(* IEC 61131-3 sources: plc-st-coding-agent/progress/evidence/f14_p1_20261111b/jobs/custom_minimax-m27, 44 files *)

(* ---- public-hard-01.candidate_01.st ---- *)
(* Material Proportioning Process Control *)
(* PLC Program in Structured Text (ST) *)

TYPE ProcessState :
    (
        IDLE        := 0,
        FILL_A      := 1,
        FILL_B      := 2,
        FILL_C      := 3,
        MIXING      := 4,
        DISCHARGE   := 5
    );
END_TYPE

VAR
    (* Internal state variables *)
    autoState         : ProcessState := IDLE;
    prevAutoStart     : BOOL := FALSE;
    prevValveAStart   : BOOL := FALSE;
    prevValveBStart   : BOOL := FALSE;
    prevValveCStart   : BOOL := FALSE;
    prevValveDStart   : BOOL := FALSE;
    prevMixMotorStart : BOOL := FALSE;
END_VAR

(* Emergency Stop - Highest Priority *)
IF NOT estop THEN
    valveARun    := FALSE;
    valveBRun    := FALSE;
    valveCRun    := FALSE;
    valveDRun    := FALSE;
    mixMotorRun  := FALSE;
    autoState    := IDLE;
    RETURN;
END_IF

(* Rising edge detection for buttons *)
IF autoStart AND NOT prevAutoStart THEN
    (* Rising edge detected for autoStart *)
END_IF

IF valveAStart AND NOT prevValveAStart THEN
    valveARun := NOT valveARun;
END_IF;

IF valveBStart AND NOT prevValveBStart THEN
    valveBRun := NOT valveBRun;
END_IF;

IF valveCStart AND NOT prevValveCStart THEN
    valveCRun := NOT valveCRun;
END_IF;

IF valveDStart AND NOT prevValveDStart THEN
    valveDRun := NOT valveDRun;
END_IF;

IF mixMotorStart AND NOT prevMixMotorStart THEN
    mixMotorRun := NOT mixMotorRun;
END_IF;

(* Update previous button states *)
prevAutoStart     := autoStart;
prevValveAStart   := valveAStart;
prevValveBStart   := valveBStart;
prevValveCStart   := valveCStart;
prevValveDStart   := valveDStart;
prevMixMotorStart := mixMotorStart;

(* Mode Selection *)
IF opeMode THEN
    (* ========== AUTOMATIC MODE ========== *)

    (* Initialize outputs to FALSE *)
    valveARun   := FALSE;
    valveBRun   := FALSE;
    valveCRun   := FALSE;
    valveDRun   := FALSE;
    mixMotorRun := FALSE;

    (* Start automatic process on rising edge of autoStart *)
    IF autoStart AND NOT prevAutoStart THEN
        IF autoState = IDLE THEN
            autoState := FILL_A;
            valveARun := TRUE;
        END_IF
    END_IF

    (* State Machine - Sequential Control *)
    IF autoState = FILL_A THEN
        valveARun := TRUE;
        (* When level reaches 50cm, close valve A and open valve B *)
        IF levelSensor >= 50 THEN
            autoState  := FILL_B;
            valveARun  := FALSE;
            valveBRun  := TRUE;
        END_IF

    ELSIF autoState = FILL_B THEN
        valveBRun := TRUE;
        (* When level reaches 80cm, close valve B *)
        IF levelSensor >= 80 THEN
            valveBRun := FALSE;

            (* Check processMode for next step *)
            IF NOT processMode THEN
                (* processMode=false: Direct to mixing *)
                autoState  := MIXING;
                mixMotorRun := TRUE;
            ELSE
                (* processMode=true: Fill material C first *)
                autoState := FILL_C;
            END_IF
        END_IF

    ELSIF autoState = FILL_C THEN
        valveCRun := TRUE;
        (* When level reaches 100cm, close valve C and start mixing *)
        IF levelSensor >= 100 THEN
            autoState  := MIXING;
            valveCRun  := FALSE;
            mixMotorRun := TRUE;
        END_IF

    ELSIF autoState = MIXING THEN
        mixMotorRun := TRUE;
        (* When mixing complete signal received, stop motor *)
        IF mixMotorComplete THEN
            autoState  := DISCHARGE;
            mixMotorRun := FALSE;
        END_IF

    ELSIF autoState = DISCHARGE THEN
        valveDRun := TRUE;
        (* After discharge, return to idle - process complete *)
        autoState := IDLE;

    END_IF

ELSE
    (* ========== MANUAL MODE ========== *)
    (* In manual mode, automatic state machine is reset *)
    autoState := IDLE;

END_IF

(* ---- public-medium-05.candidate_01.st ---- *)
// Automated Production Line Control - ST Implementation

// Define the states for automatic mode
TYPE ProductionState :
(
    WAIT_A           := 0,  // Waiting for product at Workstation A
    WAIT_A_PRESSED   := 1,  // Product at A, waiting for ButtonA press
    MOVING_AB        := 2,  // Motor moving product from A to B
    WAIT_B_PRESSED   := 3,  // Product at B, waiting for ButtonB press
    MOVING_BC        := 4,  // Motor moving product from B to C
    WAIT_C_PRESSED   := 5,  // Product at C, waiting for ButtonC press
    COMPLETE         := 6   // Product processing complete
);
END_TYPE

VAR
    // State variable for automatic mode
    State : ProductionState := WAIT_A;

    // Edge detection variables
    SensorA_Edge  : BOOL := FALSE;
    SensorB_Edge  : BOOL := FALSE;
    SensorC_Edge  : BOOL := FALSE;
    SensorA_Prev  : BOOL := FALSE;
    SensorB_Prev  : BOOL := FALSE;
    SensorC_Prev  : BOOL := FALSE;
END_VAR

// Edge detection for sensors
SensorA_Edge := SensorA AND NOT SensorA_Prev;
SensorB_Edge := SensorB AND NOT SensorB_Prev;
SensorC_Edge := SensorC AND NOT SensorC_Prev;

// Store previous sensor states for edge detection
SensorA_Prev := SensorA;
SensorB_Prev := SensorB;
SensorC_Prev := SensorC;

// Manual Mode (Mode = 0)
IF Mode = FALSE THEN
    // Reset state to initial when switching to manual mode
    State := WAIT_A;

    // Forward and reverse rotation with interlock
    // Both cannot be active at the same time
    MotorForward := ForwardButton AND NOT ReverseButton;
    MotorReverse := ReverseButton AND NOT ForwardButton;

    // Completion light is off in manual mode
    CompletionLight := FALSE;

// Automatic Mode (Mode = 1)
ELSE
    // State machine logic
    CASE State OF
        // State 0: Waiting for product at Workstation A
        WAIT_A:
            MotorForward := FALSE;
            MotorReverse := FALSE;

            // Detect product arrival at A
            IF SensorA_Edge THEN
                State := WAIT_A_PRESSED;
            END_IF

        // State 1: Product at A, waiting for operator to press ButtonA
        WAIT_A_PRESSED:
            MotorForward := FALSE;
            MotorReverse := FALSE;

            // Operator presses ButtonA to signal processing complete
            IF ButtonA THEN
                State := MOVING_AB;
            END_IF

            // Safety: If product leaves A unexpectedly, return to WAIT_A
            IF NOT SensorA THEN
                State := WAIT_A;
            END_IF

        // State 2: Motor moving product from A to B
        MOVING_AB:
            MotorForward := TRUE;
            MotorReverse := FALSE;

            // Product arrives at B
            IF SensorB THEN
                State := WAIT_B_PRESSED;
            END_IF

        // State 3: Product at B, waiting for operator to press ButtonB
        WAIT_B_PRESSED:
            MotorForward := FALSE;
            MotorReverse := FALSE;

            // Operator presses ButtonB to signal processing complete
            IF ButtonB THEN
                State := MOVING_BC;
            END_IF

            // Safety: If product leaves B unexpectedly, return to WAIT_A
            IF NOT SensorB THEN
                State := WAIT_A;
            END_IF

        // State 4: Motor moving product from B to C
        MOVING_BC:
            MotorForward := TRUE;
            MotorReverse := FALSE;

            // Product arrives at C
            IF SensorC THEN
                State := WAIT_C_PRESSED;
            END_IF

        // State 5: Product at C, waiting for operator to press ButtonC
        WAIT_C_PRESSED:
            MotorForward := FALSE;
            MotorReverse := FALSE;

            // Operator presses ButtonC to signal processing complete
            IF ButtonC THEN
                State := COMPLETE;
            END_IF

            // Safety: If product leaves C unexpectedly, return to WAIT_A
            IF NOT SensorC THEN
                State := WAIT_A;
            END_IF

        // State 6: Product processing complete
        COMPLETE:
            MotorForward := FALSE;
            MotorReverse := FALSE;

            // When product is taken away (SensorC no longer detects product)
            IF NOT SensorC THEN
                State := WAIT_A;
            END_IF

    END_CASE;

    // Set CompletionLight based on current state
    // Light is ON when product is at C and processing is complete (button pressed)
    CompletionLight := (State = COMPLETE);

END_IF;

(* ---- public-easy-02.candidate_01.st ---- *)
FUNCTION_BLOCK FB_DualWordEdgeDetection
VAR_OUTPUT
    hasChanged      : BOOL;
    hasRisingEdges  : BOOL;
    risingBits      : DWORD;
    noOfRisingBits  : USINT;
    hasFallingEdges : BOOL;
    fallingBits     : DWORD;
    noOfFallingBits : USINT;
END_VAR

VAR_INPUT
    value : DWORD;
END_VAR

VAR
    prevValue : DWORD;
END_VAR

// ============================================================================
// Internal Function: Count the number of set bits in a DWORD
// Uses Brian Kernighan's algorithm for efficiency
// ============================================================================
FUNCTION PRIVATE FB_CountBits : USINT
VAR_INPUT
    bits : DWORD;
END_VAR
VAR
    count : USINT := 0;
END_VAR
    WHILE bits <> 0 DO
        bits := bits & (bits - 1);
        count := count + 1;
    END_WHILE
    FB_CountBits := count;
END_FUNCTION

// ============================================================================
// Main Edge Detection Logic
// ============================================================================

// Rising edge detection: current = 1 AND previous = 0
risingBits := value AND (NOT prevValue);

// Falling edge detection: current = 0 AND previous = 1
fallingBits := (NOT value) AND prevValue;

// Check if the entire value has changed
hasChanged := (value <> prevValue);

// Set boolean flags for edge detection
hasRisingEdges  := (risingBits <> 16#00000000);
hasFallingEdges := (fallingBits <> 16#00000000);

// Count the number of set bits (edges) in each pattern
noOfRisingBits  := FB_CountBits(risingBits);
noOfFallingBits := FB_CountBits(fallingBits);

// Store current value for next cycle edge detection
prevValue := value;

END_FUNCTION_BLOCK

(* ---- public-easy-02.candidate_02.st ---- *)
FUNCTION_BLOCK FB_DualWordEdgeDetection
VAR
    prevValue   : DWORD;
    bitCounter  : DWORD;
    countRising : USINT;
    countFalling: USINT;
END_VAR

VAR_INPUT
    value : DWORD;
END_VAR

VAR_OUTPUT
    hasChanged      : BOOL;
    hasRisingEdges  : BOOL;
    risingBits      : DWORD;
    noOfRisingBits  : USINT;
    hasFallingEdges : BOOL;
    fallingBits     : DWORD;
    noOfFallingBits : USINT;
END_VAR

// ============================================================================
// Rising edge detection: current = 1 AND previous = 0
risingBits := value AND (NOT prevValue);

// Falling edge detection: current = 0 AND previous = 1
fallingBits := (NOT value) AND prevValue;

// Check if the entire value has changed
hasChanged := (value <> prevValue);

// Set boolean flags for edge detection
hasRisingEdges  := (risingBits <> 16#00000000);
hasFallingEdges := (fallingBits <> 16#00000000);

// ============================================================================
// Count rising edges using Brian Kernighan's algorithm
// ============================================================================
bitCounter  := risingBits;
countRising := 0;
WHILE bitCounter <> 0 DO
    bitCounter := bitCounter & (bitCounter - 1);
    countRising := countRising + 1;
END_WHILE
noOfRisingBits := countRising;

// ============================================================================
// Count falling edges using Brian Kernighan's algorithm
// ============================================================================
bitCounter   := fallingBits;
countFalling := 0;
WHILE bitCounter <> 0 DO
    bitCounter := bitCounter & (bitCounter - 1);
    countFalling := countFalling + 1;
END_WHILE
noOfFallingBits := countFalling;

// ============================================================================
// Store current value for next cycle edge detection
// ============================================================================
prevValue := value;

END_FUNCTION_BLOCK

(* ---- public-easy-03.candidate_01.st ---- *)
FUNCTION_BLOCK AlarmHyst
VAR_INPUT
    Value      : REAL;   (* Current measured value *)
    hiLevel    : REAL;   (* High‑limit alarm threshold *)
    loLevel    : REAL;   (* Low‑limit alarm threshold  *)
    hystWindow : REAL;   (* Hysteresis window width    *)
END_VAR

VAR_OUTPUT
    hiAlarm : BOOL;   (* High‑limit alarm status *)
    loAlarm : BOOL;   (* Low‑limit alarm status  *)
    error   : BOOL;   (* FALSE = normal operation, TRUE = error detected *)
    status  : WORD;   (* Status / error code (0 = OK) *)
END_VAR

(* ---------------------------------------------------------------- *)
(*  Error detection (must be performed before any alarm logic)      *)
(* ---------------------------------------------------------------- *)
IF loLevel >= hiLevel THEN
    error   := TRUE;
    status  := WORD#16#8001;           (* 16#8001 : loLevel not lower than hiLevel *)
    hiAlarm := FALSE;
    loAlarm := FALSE;
    RETURN;                            (* leave the function block *)
END_IF

IF hystWindow >= (hiLevel - loLevel) THEN
    error   := TRUE;
    status  := WORD#16#8002;           (* 16#8002 : hystWindow too large *)
    hiAlarm := FALSE;
    loAlarm := FALSE;
    RETURN;
END_IF

(* ---------------------------------------------------------------- *)
(*  Normal operation – clear error flag and execute alarm logic     *)
(* ---------------------------------------------------------------- *)
error  := FALSE;
status := WORD#0;

(* ----- High‑limit alarm with hysteresis ------------------------- *)
(* Trigger:   Value > hiLevel                                       *)
(* Clear:     Value < hiLevel - hystWindow                          *)
IF Value > hiLevel THEN
    hiAlarm := TRUE;
ELSIF Value < (hiLevel - hystWindow) THEN
    hiAlarm := FALSE;
END_IF

(* ----- Low‑limit alarm with hysteresis -------------------------- *)
(* Trigger:   Value < loLevel                                       *)
(* Clear:     Value > loLevel + hystWindow                          *)
IF Value < loLevel THEN
    loAlarm := TRUE;
ELSIF Value > (loLevel + hystWindow) THEN
    loAlarm := FALSE;
END_IF

END_FUNCTION_BLOCK

(* ---- public-easy-03.candidate_02.st ---- *)
FUNCTION_BLOCK AlarmHyst
VAR_INPUT
    Value      : REAL;
    hiLevel    : REAL;
    loLevel    : REAL;
    hystWindow : REAL;
END_VAR

VAR_OUTPUT
    hiAlarm : BOOL;
    loAlarm : BOOL;
    error   : BOOL;
    status  : WORD;
END_VAR

VAR RETAIN
    errorOccurred : BOOL := FALSE;
    statusValue   : WORD := WORD#0;
    hiAlarmPrev   : BOOL := FALSE;
    loAlarmPrev   : BOOL := FALSE;
END_VAR

(* ---------------------------------------------------------------- *)
(*  Error detection - latch error state                             *)
(* ---------------------------------------------------------------- *)
IF loLevel >= hiLevel THEN
    error         := TRUE;
    status        := WORD#16#8001;
    errorOccurred := TRUE;
    statusValue   := WORD#16#8001;
    hiAlarm       := FALSE;
    loAlarm       := FALSE;
    RETURN;
END_IF

IF hystWindow >= (hiLevel - loLevel) THEN
    error         := TRUE;
    status        := WORD#16#8002;
    errorOccurred := TRUE;
    statusValue   := WORD#16#8002;
    hiAlarm       := FALSE;
    loAlarm       := FALSE;
    RETURN;
END_IF

(* ---------------------------------------------------------------- *)
(*  Normal operation                                                *)
(* ---------------------------------------------------------------- *)
(* Clear latched error when configuration is valid                  *)
errorOccurred := FALSE;
statusValue   := WORD#0;

(* ----- High‑limit alarm with hysteresis ------------------------- *)
IF Value > hiLevel THEN
    hiAlarmPrev := TRUE;
ELSIF Value < (hiLevel - hystWindow) THEN
    hiAlarmPrev := FALSE;
END_IF

(* ----- Low‑limit alarm with hysteresis -------------------------- *)
IF Value < loLevel THEN
    loAlarmPrev := TRUE;
ELSIF Value > (loLevel + hystWindow) THEN
    loAlarmPrev := FALSE;
END_IF

(* Update outputs *)
error   := errorOccurred;
status  := statusValue;
hiAlarm := hiAlarmPrev;
loAlarm := loAlarmPrev;

END_FUNCTION_BLOCK

(* ---- public-easy-04.candidate_01.st ---- *)
(* -------------------------------------------------------------
   Jam Pump Debouncing and Runtime Maintenance
   -------------------------------------------------------------
   Inputs
      VISCOSITY_OK    : Raw viscosity‑OK signal (TRUE = within range)
      PASTE_E_STOP_NC : Emergency‑stop circuit, normally closed
      DebounceTime    : Required ON‑time for the viscosity signal
      CycleTime       : Actual invocation interval (must be >0)

   Outputs
      VFD_RUN         : VFD run command (TRUE = allowed)
      PUMP_MAINT_DUE  : Maintenance‑due flag (TRUE after 500 h run)
      PUMP_RUNTIME_ACC: Accumulated run time (LTIME)

   Internal variables
      viscosity_valid : Viscosity condition accepted after debounce
      DebounceTimer   : TON used for debouncing
      prevEStop       : Previous state of PASTE_E_STOP_NC (edge detection)
      init            : Power‑up initialisation flag
   ------------------------------------------------------------- *)
FUNCTION_BLOCK JamPumpControl
VAR_INPUT
    VISCOSITY_OK    : BOOL;
    PASTE_E_STOP_NC : BOOL;
    DebounceTime    : TIME;
    CycleTime       : TIME;
END_VAR
VAR_OUTPUT
    VFD_RUN         : BOOL;
    PUMP_MAINT_DUE  : BOOL;
    PUMP_RUNTIME_ACC: LTIME;
END_VAR
VAR
    viscosity_valid : BOOL := FALSE;
    DebounceTimer   : TON;
    prevEStop       : BOOL := TRUE;   // assume not in emergency stop at start‑up
    init            : BOOL := TRUE;   // power‑up initialization flag
END_VAR

// -------------------------------------------------------------------
// Power‑up initialisation
// -------------------------------------------------------------------
IF init THEN
    VFD_RUN          := FALSE;            // run output OFF
    PUMP_RUNTIME_ACC := LTIME#0;         // accumulated time = 0
    PUMP_MAINT_DUE   := FALSE;           // maintenance flag cleared
    viscosity_valid  := FALSE;           // no valid viscosity yet
    DebounceTimer(IN := FALSE, PT := DebounceTime); // timer reset
    // Initialise previous E‑Stop state to current value so that a
    // spurious falling‑edge is not generated on the first scan.
    prevEStop := PASTE_E_STOP_NC;
    init := FALSE;

// -------------------------------------------------------------------
// Normal (cyclic) processing
// -------------------------------------------------------------------
ELSE

    // ---- Emergency‑stop edge detection --------------------------------
    // If the emergency‑stop circuit opens (falling edge) the viscosity
    // permissive must be cleared and any in‑progress debounce aborted.
    IF (NOT PASTE_E_STOP_NC) AND prevEStop THEN
        viscosity_valid      := FALSE;
        DebounceTimer(IN := FALSE);   // abort timer
    END_IF
    prevEStop := PASTE_E_STOP_NC;

    // ---- Viscosity signal – immediate invalidation --------------------
    IF NOT VISCOSITY_OK THEN
        viscosity_valid := FALSE;   // loss of signal → invalid immediately
    END_IF

    // ---- Debounce timer ------------------------------------------------
    // Start timing only when:
    //   • raw signal is TRUE,
    //   • we do not yet have a valid reading,
    //   • emergency‑stop circuit is closed.
    DebounceTimer(
        IN := VISCOSITY_OK AND NOT viscosity_valid AND PASTE_E_STOP_NC,
        PT := DebounceTime
    );
    DebounceTimer();   // execute the TON block

    // When the timer finishes, the viscosity condition becomes valid.
    IF DebounceTimer.Q THEN
        viscosity_valid := TRUE;
    END_IF

    // ---- Run permissive ------------------------------------------------
    // VFD may run only when the emergency‑stop is closed AND the
    // viscosity condition has been accepted after debounce.
    VFD_RUN := PASTE_E_STOP_NC AND viscosity_valid;

    // ---- Runtime accumulation -----------------------------------------
    // Accumulate time only while the pump is actually running.
    IF VFD_RUN THEN
        PUMP_RUNTIME_ACC := PUMP_RUNTIME_ACC + LTIME(CycleTime);
    END_IF

    // ---- Maintenance‑due indication ------------------------------------
    // Informational flag – does not affect safety or operation.
    PUMP_MAINT_DUE := (PUMP_RUNTIME_ACC >= LTIME#500h);

END_IF

END_FUNCTION_BLOCK

(* ---- public-easy-04.candidate_02.st ---- *)
(* -------------------------------------------------------------
   Jam Pump Debouncing and Runtime Maintenance
   -------------------------------------------------------------
   Inputs
      VISCOSITY_OK    : Raw viscosity‑OK signal (TRUE = within range)
      PASTE_E_STOP_NC : Emergency‑stop circuit, normally closed
      DebounceTime    : Required ON‑time for the viscosity signal
      CycleTime       : Actual invocation interval (must be >0)

   Outputs
      VFD_RUN         : VFD run command (TRUE = allowed)
      PUMP_MAINT_DUE  : Maintenance‑due flag (TRUE after 500 h run)
      PUMP_RUNTIME_ACC: Accumulated run time (LTIME)

   Internal variables
      viscosity_valid : Viscosity condition accepted after debounce
      DebounceTimer   : TON used for debouncing
      prevEStop       : Previous state of PASTE_E_STOP_NC (edge detection)
      init            : Power‑up initialisation flag
   ------------------------------------------------------------- *)
FUNCTION_BLOCK JamPumpControl
VAR_INPUT
    VISCOSITY_OK    : BOOL;
    PASTE_E_STOP_NC : BOOL;
    DebounceTime    : TIME;
    CycleTime       : TIME;
END_VAR
VAR_OUTPUT
    VFD_RUN         : BOOL;
    PUMP_MAINT_DUE  : BOOL;
    PUMP_RUNTIME_ACC: LTIME;
END_VAR
VAR
    viscosity_valid : BOOL := FALSE;
    DebounceTimer   : TON;
    prevEStop       : BOOL := TRUE;   // assume not in emergency stop at start‑up
    init            : BOOL := TRUE;   // power‑up initialization flag
END_VAR

// -------------------------------------------------------------------
// Power‑up initialisation
// -------------------------------------------------------------------
IF init THEN
    VFD_RUN          := FALSE;            // run output OFF
    PUMP_RUNTIME_ACC := LTIME#0h;        // accumulated time = 0
    PUMP_MAINT_DUE   := FALSE;           // maintenance flag cleared
    viscosity_valid  := FALSE;           // no valid viscosity yet
    DebounceTimer(IN := FALSE, PT := DebounceTime); // timer reset
    // Initialise previous E‑Stop state to current value so that a
    // spurious falling‑edge is not generated on the first scan.
    prevEStop := PASTE_E_STOP_NC;
    init := FALSE;

// -------------------------------------------------------------------
// Normal (cyclic) processing
// -------------------------------------------------------------------
ELSE

    // ---- Emergency‑stop edge detection --------------------------------
    // If the emergency‑stop circuit opens (falling edge) the viscosity
    // permissive must be cleared and any in‑progress debounce aborted.
    IF (NOT PASTE_E_STOP_NC) AND prevEStop THEN
        viscosity_valid      := FALSE;
        DebounceTimer(IN := FALSE);   // abort timer
    END_IF
    prevEStop := PASTE_E_STOP_NC;

    // ---- Viscosity signal – immediate invalidation --------------------
    IF NOT VISCOSITY_OK THEN
        viscosity_valid := FALSE;   // loss of signal → invalid immediately
    END_IF

    // ---- Debounce timer ------------------------------------------------
    // Start timing only when:
    //   • raw signal is TRUE,
    //   • we do not yet have a valid reading,
    //   • emergency‑stop circuit is closed.
    DebounceTimer(
        IN := VISCOSITY_OK AND NOT viscosity_valid AND PASTE_E_STOP_NC,
        PT := DebounceTime
    );
    DebounceTimer();   // execute the TON block

    // When the timer finishes, the viscosity condition becomes valid.
    IF DebounceTimer.Q THEN
        viscosity_valid := TRUE;
    END_IF

    // ---- Run permissive ------------------------------------------------
    // VFD may run only when the emergency‑stop is closed AND the
    // viscosity condition has been accepted after debounce.
    VFD_RUN := PASTE_E_STOP_NC AND viscosity_valid;

    // ---- Runtime accumulation -----------------------------------------
    // Accumulate time only while the pump is actually running.
    // TIME values implicitly convert to LTIME in expressions.
    IF VFD_RUN THEN
        PUMP_RUNTIME_ACC := PUMP_RUNTIME_ACC + CycleTime;
    END_IF

    // ---- Maintenance‑due indication ------------------------------------
    // Informational flag – does not affect safety or operation.
    PUMP_MAINT_DUE := (PUMP_RUNTIME_ACC >= LTIME#500h);

END_IF

END_FUNCTION_BLOCK

(* ---- public-hard-03.candidate_02.st ---- *)
FUNCTION_BLOCK RecipeManagement
VAR_INPUT
    addRecipe    : BOOL;
    deleteRecipe : BOOL;
    modifyRecipe : BOOL;
    queryRecipe  : BOOL;
    recipeIn     : ST_Recipe;
END_VAR

VAR_OUTPUT
    recipeAdded       : BOOL;
    recipeDeleted     : BOOL;
    recipeModified    : BOOL;
    recipeQueryResult : ST_Recipe;
    error             : BOOL;
    status            : WORD;
END_VAR

VAR_IN_OUT
    recipe : ARRAY[1..10] OF ST_Recipe;
END_VAR

VAR
    i              : INT;
    foundIndex     : INT;
    emptySlotIndex : INT;
    found          : BOOL;
END_VAR

//---------------------------------------------------------------------------
// Initialization
//---------------------------------------------------------------------------
error            := FALSE;
status           := 16#0000;
recipeAdded      := FALSE;
recipeDeleted    := FALSE;
recipeModified   := FALSE;
recipeQueryResult.recipeID              := 0;
recipeQueryResult.ingredientType        := 0;
recipeQueryResult.ingredientRatio       := 0.0;
recipeQueryResult.productionTemperature := 0.0;

//---------------------------------------------------------------------------
// Query Recipe Operation
//---------------------------------------------------------------------------
IF queryRecipe THEN
    found      := FALSE;
    foundIndex := 0;

    FOR i := 1 TO 10 DO
        IF recipe[i].recipeID = recipeIn.recipeID THEN
            found      := TRUE;
            foundIndex := i;
            EXIT;
        END_IF
    END_FOR

    IF found THEN
        recipeQueryResult := recipe[foundIndex];
        error  := FALSE;
        status := 16#0000;
    ELSE
        error  := TRUE;
        status := 16#8001;
    END_IF
END_IF

//---------------------------------------------------------------------------
// Add Recipe Operation
//---------------------------------------------------------------------------
IF addRecipe THEN
    found      := FALSE;
    foundIndex := 0;

    // Check for duplicate recipeID
    FOR i := 1 TO 10 DO
        IF recipe[i].recipeID = recipeIn.recipeID THEN
            found := TRUE;
            EXIT;
        END_IF
    END_FOR

    IF found THEN
        error  := TRUE;
        status := 16#8002;
    ELSE
        // Find first empty slot (smallest index)
        found          := FALSE;
        emptySlotIndex := 0;

        FOR i := 1 TO 10 DO
            IF recipe[i].recipeID = 0 THEN
                emptySlotIndex := i;
                found          := TRUE;
                EXIT;
            END_IF
        END_FOR

        IF NOT found THEN
            error  := TRUE;
            status := 16#8003;
        ELSE
            recipe[emptySlotIndex] := recipeIn;
            recipeAdded            := TRUE;
            error                  := FALSE;
            status                 := 16#0000;
        END_IF
    END_IF
END_IF

//---------------------------------------------------------------------------
// Delete Recipe Operation
//---------------------------------------------------------------------------
IF deleteRecipe THEN
    found      := FALSE;
    foundIndex := 0;

    FOR i := 1 TO 10 DO
        IF recipe[i].recipeID = recipeIn.recipeID THEN
            found      := TRUE;
            foundIndex := i;
            EXIT;
        END_IF
    END_FOR

    IF found THEN
        recipe[foundIndex].recipeID              := 0;
        recipe[foundIndex].ingredientType        := 0;
        recipe[foundIndex].ingredientRatio       := 0.0;
        recipe[foundIndex].productionTemperature := 0.0;
        recipeDeleted                            := TRUE;
        error                                    := FALSE;
        status                                   := 16#0000;
    ELSE
        error  := TRUE;
        status := 16#8004;
    END_IF
END_IF

//---------------------------------------------------------------------------
// Modify Recipe Operation
//---------------------------------------------------------------------------
IF modifyRecipe THEN
    found      := FALSE;
    foundIndex := 0;

    FOR i := 1 TO 10 DO
        IF recipe[i].recipeID = recipeIn.recipeID THEN
            found      := TRUE;
            foundIndex := i;
            EXIT;
        END_IF
    END_FOR

    IF found THEN
        recipe[foundIndex] := recipeIn;
        recipeModified     := TRUE;
        error              := FALSE;
        status             := 16#0000;
    ELSE
        error  := TRUE;
        status := 16#8005;
    END_IF
END_IF

END_FUNCTION_BLOCK

(* ---- public-hard-04.candidate_01.st ---- *)
(* --------------------------------------------------
   FUNCTION BLOCK FIFO
   First‑In‑First‑Out circular queue using the caller‑supplied buffer.
   Derives capacity and element type from the buffer.
   -------------------------------------------------- *)
FUNCTION_BLOCK FIFO
VAR_INPUT
    enqueue  : BOOL;      (* Rising edge → enqueue one item           *)
    dequeue  : BOOL;      (* Rising edge → dequeue one item           *)
    reset    : BOOL;      (* TRUE → empty the queue, highest priority *)
END_VAR
VAR_OUTPUT
    elementCount : DINT;  (* Number of valid elements (0 … capacity) *)
    status       : WORD;  (* 16#0000, 16#8001, 16#8002                *)
END_VAR
VAR_IN_OUT
    item   : VARIANT;     (* Scalar to read (enqueue) or write (dequeue) *)
    buffer : VARIANT;     (* One‑dimensional array used as storage       *)
END_VAR

VAR
    (* Internal queue state --------------------------------------------------- *)
    headIndex   : DINT;   (* Current head position (real array index)        *)
    tailIndex   : DINT;   (* Current tail position (real array index)        *)
    count       : DINT;   (* Number of stored elements (mirrors elementCount) *)

    (* Array bounds (re‑computed each cycle because buffer never changes) ----- *)
    lowerBound  : DINT;   (* LOWER_BOUND(buffer,1)                           *)
    upperBound  : DINT;   (* UPPER_BOUND(buffer,1)                           *)
    capacity    : DINT;   (* upperBound - lowerBound + 1                     *)

    (* Edge detection --------------------------------------------------------- *)
    prevEnqueue : BOOL;   (* Value of enqueue from previous cycle            *)
    prevDequeue : BOOL;   (* Value of dequeue from previous cycle            *)
    enqueueRising : BOOL; (* TRUE on a rising edge of enqueue                *)
    dequeueRising : BOOL; (* TRUE on a rising edge of dequeue                *)

    (* First‑call initialization ---------------------------------------------- *)
    initDone    : BOOL;   (* TRUE after the first execution                  *)
END_VAR

(* -------------------------------------------------------------------------- *)
(* Body of the function block                                                 *)
(* -------------------------------------------------------------------------- *)

(* 1. Determine capacity from the supplied buffer ----------------------------- *)
lowerBound := LOWER_BOUND(buffer, 1);
upperBound := UPPER_BOUND(buffer, 1);
capacity   := upperBound - lowerBound + 1;

(* 2. Initialise internal variables on the very first call ------------------- *)
IF NOT initDone THEN
    headIndex := lowerBound;
    tailIndex := lowerBound;
    count     := 0;
    initDone  := TRUE;
END_IF

(* 3. Reset handling (highest priority) ------------------------------------- *)
IF reset THEN
    count     := 0;
    headIndex := lowerBound;
    tailIndex := lowerBound;
    status    := 16#0000;                     (* no error                     *)
ELSE
    (* 4. Detect rising edges on enqueue / dequeue --------------------------- *)
    enqueueRising := enqueue AND NOT prevEnqueue;
    dequeueRising := dequeue AND NOT prevDequeue;

    (* Store current input states for next cycle ----------------------------- *)
    prevEnqueue := enqueue;
    prevDequeue := dequeue;

    (* Default status = no error -------------------------------------------- *)
    status := 16#0000;

    (* 5. Enqueue request ----------------------------------------------------- *)
    IF enqueueRising THEN
        IF count < capacity THEN
            (* Append the current item to the tail -------------------------- *)
            buffer[tailIndex] := item;

            (* Advance tail (circular) -------------------------------------- *)
            tailIndex := tailIndex + 1;
            IF tailIndex > upperBound THEN
                tailIndex := lowerBound;
            END_IF

            count := count + 1;
        ELSE
            (* Queue full – reject the request -------------------------------- *)
            status := 16#8002;
        END_IF
    END_IF

    (* 6. Dequeue request ----------------------------------------------------- *)
    IF dequeueRising THEN
        IF count > 0 THEN
            (* Copy the front element to item -------------------------------- *)
            item := buffer[headIndex];

            (* Advance head (circular) --------------------------------------- *)
            headIndex := headIndex + 1;
            IF headIndex > upperBound THEN
                headIndex := lowerBound;
            END_IF

            count := count - 1;
        ELSE
            (* Queue empty – reject the request ------------------------------- *)
            status := 16#8001;
        END_IF
    END_IF
END_IF

(* 7. Publish the current number of stored elements -------------------------- *)
elementCount := count;

END_FUNCTION_BLOCK

(* ---- public-hard-06.candidate_02.st ---- *)
FUNCTION_BLOCK ProductionControl
VAR_INPUT
    Mode            : BOOL;          (* 0 = Manual, 1 = Automatic *)
    ForwardButton   : BOOL;          (* Manual forward command *)
    ReverseButton   : BOOL;          (* Manual reverse command *)
    SensorFeed      : BOOL;          (* Material at loading station *)
    SensorWash      : BOOL;          (* Material at cleaning station *)
    SensorWeight    : BOOL;          (* Material at weighing station *)
    SensorFiring    : BOOL;          (* Product at firing station *)
    SensorOutput    : BOOL;          (* Product at finished-product station *)
    washComplete    : BOOL;          (* Cleaning finished *)
    weightComplete  : BOOL;          (* Weighing finished *)
    weight          : REAL;          (* Measured weight *)
    firingComplete  : BOOL;          (* Firing finished *)
END_VAR

VAR_OUTPUT
    MotorForward    : BOOL;          (* Motor forward rotation *)
    MotorReverse    : BOOL;          (* Motor reverse rotation *)
    kick            : BOOL;          (* Rejection command *)
    CompletionLight : BOOL;          (* Product ready light *)
    firingTemp      : REAL;          (* Calculated firing temperature *)
END_VAR

VAR
    curState        : INT := 0;      (* Current automatic state *)
    lastSensorFeed    : BOOL := FALSE;
    lastSensorWash    : BOOL := FALSE;
    lastSensorWeight  : BOOL := FALSE;
    lastSensorFiring  : BOOL := FALSE;
    lastSensorOutput  : BOOL := FALSE;
    lastWashComplete  : BOOL := FALSE;
    lastWeightComplete: BOOL := FALSE;
    lastFiringComplete: BOOL := FALSE;
    sensorFeedRising    : BOOL;
    sensorWashRising    : BOOL;
    sensorWeightRising  : BOOL;
    sensorFiringRising  : BOOL;
    sensorOutputRising  : BOOL;
    sensorOutputFalling : BOOL;
    washCompleteRising  : BOOL;
    weightCompleteRising: BOOL;
    firingCompleteRising: BOOL;
    washProcessed   : BOOL := FALSE;
    weightProcessed : BOOL := FALSE;
    firingProcessed : BOOL := FALSE;
END_VAR

(* Edge detection *)
sensorFeedRising     := SensorFeed     AND NOT lastSensorFeed;
sensorWashRising     := SensorWash     AND NOT lastSensorWash;
sensorWeightRising   := SensorWeight   AND NOT lastSensorWeight;
sensorFiringRising   := SensorFiring   AND NOT lastSensorFiring;
sensorOutputRising   := SensorOutput   AND NOT lastSensorOutput;
sensorOutputFalling  := NOT SensorOutput AND lastSensorOutput;
washCompleteRising   := washComplete   AND NOT lastWashComplete;
weightCompleteRising := weightComplete AND NOT lastWeightComplete;
firingCompleteRising := firingComplete AND NOT lastFiringComplete;

lastSensorFeed     := SensorFeed;
lastSensorWash     := SensorWash;
lastSensorWeight   := SensorWeight;
lastSensorFiring   := SensorFiring;
lastSensorOutput   := SensorOutput;
lastWashComplete   := washComplete;
lastWeightComplete := weightComplete;
lastFiringComplete := firingComplete;

(* Mode handling *)
IF Mode = FALSE THEN
    MotorForward    := FALSE;
    MotorReverse    := FALSE;
    kick            := FALSE;
    CompletionLight := FALSE;
    firingTemp      := 0.0;
    curState        := 0;
    washProcessed   := FALSE;
    weightProcessed := FALSE;
    firingProcessed := FALSE;

    IF ForwardButton AND NOT ReverseButton THEN
        MotorForward := TRUE;
    ELSE
        MotorForward := FALSE;
    END_IF

    IF ReverseButton AND NOT ForwardButton THEN
        MotorReverse := TRUE;
    ELSE
        MotorReverse := FALSE;
    END_IF
ELSE
    MotorReverse := FALSE;

    CASE curState OF
        0: (* IDLE *)
            IF sensorFeedRising THEN
                curState     := 1;
                MotorForward := TRUE;
            ELSE
                MotorForward    := FALSE;
                kick            := FALSE;
                CompletionLight := FALSE;
                firingTemp      := 0.0;
            END_IF

        1: (* MOVING_TO_WASH *)
            IF sensorWashRising THEN
                MotorForward := FALSE;
                curState     := 2;
                washProcessed := FALSE;
            END_IF

        2: (* AT_WASH *)
            IF washCompleteRising AND NOT washProcessed THEN
                MotorForward := TRUE;
                curState      := 3;
                washProcessed := TRUE;
            END_IF

        3: (* MOVING_TO_WEIGH *)
            IF sensorWeightRising THEN
                MotorForward    := FALSE;
                curState        := 4;
                weightProcessed := FALSE;
            END_IF

        4: (* AT_WEIGH *)
            IF weightCompleteRising AND NOT weightProcessed THEN
                weightProcessed := TRUE;
                IF weight >= 100.0 AND weight <= 200.0 THEN
                    firingTemp  := 500.0 + ((weight - 100.0) / 100.0) * 50.0;
                    MotorForward := TRUE;
                    curState     := 5;
                ELSE
                    kick         := TRUE;
                    MotorForward := FALSE;
                    curState     := 9;
                END_IF
            END_IF

        5: (* MOVING_TO_FIRING *)
            IF sensorFiringRising THEN
                MotorForward    := FALSE;
                curState        := 6;
                firingProcessed := FALSE;
            END_IF

        6: (* AT_FIRING *)
            IF firingCompleteRising AND NOT firingProcessed THEN
                MotorForward    := TRUE;
                curState         := 7;
                firingProcessed  := TRUE;
            END_IF

        7: (* MOVING_TO_OUTPUT *)
            IF sensorOutputRising THEN
                MotorForward    := FALSE;
                CompletionLight := TRUE;
                curState        := 8;
            END_IF

        8: (* AT_OUTPUT *)
            CompletionLight := SensorOutput;
            IF sensorOutputFalling THEN
                CompletionLight := FALSE;
                curState        := 0;
                firingTemp      := 0.0;
                kick            := FALSE;
            END_IF

        9: (* REJECT *)
            kick         := TRUE;
            MotorForward := FALSE;
            IF NOT SensorWeight THEN
                kick     := FALSE;
                curState := 0;
            END_IF

    END_CASE
END_IF

END_FUNCTION_BLOCK

(* ---- public-medium-01.candidate_01.st ---- *)
(*--------------------------------------------------------------
  Data‑type for a single pump
--------------------------------------------------------------*)
TYPE ST_Pump : STRUCT
    priority  : INT;     // Read‑only priority (larger → higher priority)
    selection : BOOL;    // Read‑only manual‑selection flag
    RunComd   : BOOL;    // Write‑only run command (TRUE = start, FALSE = stop)
END_STRUCT
END_TYPE

(*--------------------------------------------------------------
  Multi‑pump switching control function block

  Inputs:
    mode   – FALSE = manual mode, TRUE = automatic mode
    start  – start push‑button (rising‑edge triggered)
    stop   – stop push‑button (rising‑edge triggered)

  In‑Out:
    pumpGroup – array of 5 pump records (priority & selection are read,
                RunComd is written)
--------------------------------------------------------------*)
FUNCTION_BLOCK MultiPumpControl
VAR_INPUT
    mode  : BOOL;   // FALSE = Manual, TRUE = Automatic
    start : BOOL;   // Start push‑button (rising edge)
    stop  : BOOL;   // Stop push‑button (rising edge)
END_VAR
VAR_IN_OUT
    pumpGroup : ARRAY[1..5] OF ST_Pump;
END_VAR
VAR
    startPrev : BOOL := FALSE;   // Edge‑detection memory for START
    stopPrev  : BOOL := FALSE;   // Edge‑detection memory for STOP
    i, j, tmp : INT;             // Loop counters & temp for sorting
    sortedIdx : ARRAY[1..5] OF INT; // Indices of pumps sorted by priority
END_VAR

(* -------------------------------------------------------------
   STOP – rising edge of the STOP button stops all pumps
   ------------------------------------------------------------- *)
IF stop AND NOT stopPrev THEN
    FOR i := 1 TO 5 DO
        pumpGroup[i].RunComd := FALSE;
    END_FOR;
END_IF;
stopPrev := stop;

(* -------------------------------------------------------------
   START – rising edge of the START button starts the selected
   pump(s) in manual mode, or the three highest‑priority pumps
   in automatic mode.
   ------------------------------------------------------------- *)
IF start AND NOT startPrev THEN
    IF NOT mode THEN
        (* ---- Manual mode ---- *)
        (* Start every pump whose selection flag is TRUE *)
        FOR i := 1 TO 5 DO
            IF pumpGroup[i].selection THEN
                pumpGroup[i].RunComd := TRUE;
            END_IF;
        END_FOR;
    ELSE
        (* ---- Automatic mode ---- *)
        (* 1) Build a list of pump indices sorted by priority (descending) *)
        FOR i := 1 TO 5 DO
            sortedIdx[i] := i;
        END_FOR;

        (* Simple bubble‑sort (stable) – fine for only 5 pumps *)
        FOR i := 1 TO 4 DO
            FOR j := i+1 TO 5 DO
                IF pumpGroup[sortedIdx[j]].priority > pumpGroup[sortedIdx[i]].priority THEN
                    tmp := sortedIdx[i];
                    sortedIdx[i] := sortedIdx[j];
                    sortedIdx[j] := tmp;
                END_IF;
            END_FOR;
        END_FOR;

        (* 2) Drive the three highest‑priority pumps, keep the rest on standby *)
        FOR i := 1 TO 5 DO
            IF i <= 3 THEN
                pumpGroup[sortedIdx[i]].RunComd := TRUE;   // start
            ELSE
                pumpGroup[sortedIdx[i]].RunComd := FALSE;  // standby
            END_IF;
        END_FOR;
    END_IF;
END_IF;
startPrev := start;

END_FUNCTION_BLOCK

(* ---- public-medium-01.candidate_02.st ---- *)
(*--------------------------------------------------------------
  Data‑type for a single pump
--------------------------------------------------------------*)
TYPE ST_Pump : STRUCT
    priority  : INT;     // Read‑only priority (larger → higher priority)
    selection : BOOL;    // Read‑only manual‑selection flag
    RunComd   : BOOL;    // Write‑only run command (TRUE = start, FALSE = stop)
END_STRUCT
END_TYPE

(*--------------------------------------------------------------
  Multi‑pump switching control function block

  Inputs:
    mode   – FALSE = Manual mode, TRUE = Automatic mode
    start  – Start push‑button (rising‑edge triggered)
    stop   – Stop push‑button (rising‑edge triggered)

  In‑Out:
    pumpGroup – array of 5 pump records (priority & selection are read,
                RunComd is written)
--------------------------------------------------------------*)
FUNCTION_BLOCK MultiPumpControl
VAR_INPUT
    mode  : BOOL;   // FALSE = Manual, TRUE = Automatic
    start : BOOL;   // Start push‑button (rising edge)
    stop  : BOOL;   // Stop push‑button (rising edge)
END_VAR
VAR_IN_OUT
    pumpGroup : ARRAY[1..5] OF ST_Pump;
END_VAR
VAR
    startPrev : BOOL := FALSE;   // Edge‑detection memory for START
    stopPrev  : BOOL := FALSE;   // Edge‑detection memory for STOP
    i, j, tmp : INT;             // Loop counters & temp for sorting
    sortedIdx : ARRAY[1..5] OF INT; // Indices of pumps sorted by priority
END_VAR

(* -------------------------------------------------------------
   STOP – rising edge of the STOP button stops all pumps
   ------------------------------------------------------------- *)
IF stop AND NOT stopPrev THEN
    FOR i := 1 TO 5 DO
        pumpGroup[i].RunComd := FALSE;
    END_FOR;
END_IF;
stopPrev := stop;

(* -------------------------------------------------------------
   START – rising edge of the START button starts the selected
   pump(s) in manual mode, or the three highest‑priority pumps
   in automatic mode.
   ------------------------------------------------------------- *)
IF start AND NOT startPrev THEN
    IF NOT mode THEN
        (* ---- Manual mode ---- *)
        (* Start ONE pump: the highest‑priority pump among those selected *)
        selectedPump := 0;
        maxPriority := -1;
        FOR i := 1 TO 5 DO
            IF pumpGroup[i].selection AND pumpGroup[i].priority > maxPriority THEN
                maxPriority := pumpGroup[i].priority;
                selectedPump := i;
            END_IF;
        END_FOR;

        (* Set all pumps: selected one runs, others standby *)
        FOR i := 1 TO 5 DO
            IF i = selectedPump THEN
                pumpGroup[i].RunComd := TRUE;
            ELSE
                pumpGroup[i].RunComd := FALSE;
            END_IF;
        END_FOR;
    ELSE
        (* ---- Automatic mode ---- *)
        (* 1) Build a list of pump indices sorted by priority (descending) *)
        FOR i := 1 TO 5 DO
            sortedIdx[i] := i;
        END_FOR;

        (* Simple bubble‑sort – fine for only 5 pumps *)
        FOR i := 1 TO 4 DO
            FOR j := i+1 TO 5 DO
                IF pumpGroup[sortedIdx[j]].priority > pumpGroup[sortedIdx[i]].priority THEN
                    tmp := sortedIdx[i];
                    sortedIdx[i] := sortedIdx[j];
                    sortedIdx[j] := tmp;
                END_IF;
            END_FOR;
        END_FOR;

        (* 2) Drive the three highest‑priority pumps, keep the rest on standby *)
        FOR i := 1 TO 5 DO
            IF i <= 3 THEN
                pumpGroup[sortedIdx[i]].RunComd := TRUE;   // start (3 in use)
            ELSE
                pumpGroup[sortedIdx[i]].RunComd := FALSE;  // standby (2 on standby)
            END_IF;
        END_FOR;
    END_IF;
END_IF;
startPrev := start;

END_FUNCTION_BLOCK

(* ---- public-medium-02.candidate_01.st ---- *)
(*--------------------------------------------------------------
  Type definition for a single analog channel.
--------------------------------------------------------------*)
TYPE ST_AnalogChannel
STRUCT
    enable        : BOOL;      (* Channel conversion enable *)
    hiLIM         : REAL;      (* Upper engineering‑unit limit *)
    loLIM         : REAL;      (* Lower engineering‑unit limit *)
    bipolar       : BOOL;      (* FALSE → unipolar, TRUE → bipolar *)
    measuringMode : INT;       (* 0 = linear, 1 = std temp, 2 = climatic *)
    retVal        : WORD;      (* Per‑channel status code (output) *)
    outputValue   : REAL;      (* Converted engineering value (output) *)
END_STRUCT
END_TYPE

(*--------------------------------------------------------------
  Function block: FB_AnalogBatchProcessing
  Processes up to *count* analog channels.
--------------------------------------------------------------*)
FUNCTION_BLOCK FB_AnalogBatchProcessing
VAR_INPUT
    count : DINT;                      (* Number of channels to process *)
END_VAR
VAR_IN_OUT
    analogValues : ARRAY[*] OF INT;    (* Raw analog values (read‑only) *)
    channels     : ARRAY[*] OF ST_AnalogChannel; (* Channel settings & results *)
END_VAR
VAR
    i          : DINT;
    idxA       : INT;
    idxC       : INT;
    lowerA     : INT;
    lowerC     : INT;
    rawValue   : INT;
    rawMin     : REAL;
    rawMax     : REAL;
    scale      : REAL;
    ch         : ST_AnalogChannel;
END_VAR

    (* Determine the lower bounds of the variable‑length arrays *)
    lowerA := LOWER_BOUND(analogValues, 1);
    lowerC := LOWER_BOUND(channels, 1);

    FOR i := 0 TO count - 1 DO
        idxA := lowerA + INT#(i);
        idxC := lowerC + INT#(i);

        (* Read the channel configuration (read‑only) *)
        ch := channels[idxC];

        (* If the channel is disabled, just clear its outputs *)
        IF NOT ch.enable THEN
            channels[idxC].retVal      := 16#0000;   (* No error *)
            channels[idxC].outputValue := 0.0;
            CONTINUE;
        END_IF

        (* Read the raw analog value (read‑only) *)
        rawValue := analogValues[idxA];

        (* Branch according to measuring mode *)
        CASE ch.measuringMode OF
            0: (* ---- Non‑temperature linear scaling ---- *)
                (* Check that hiLIM > loLIM *)
                IF ch.hiLIM <= ch.loLIM THEN
                    channels[idxC].retVal      := 16#8002;  (* Range error *)
                    channels[idxC].outputValue := 0.0;
                ELSE
                    (* Determine the raw value range *)
                    IF ch.bipolar THEN
                        rawMin := -27648.0;
                        rawMax :=  27648.0;
                    ELSE
                        rawMin := 0.0;
                        rawMax := 27648.0;
                    END_IF

                    (* Linear conversion *)
                    scale := (ch.hiLIM - ch.loLIM) / (rawMax - rawMin);
                    channels[idxC].outputValue := ch.loLIM
                                 + (INT_TO_REAL(rawValue) - rawMin) * scale;
                    channels[idxC].retVal := 16#0000;      (* Success *)
                END_IF

            1: (* ---- Standard‑temperature conversion ---- *)
                channels[idxC].outputValue := INT_TO_REAL(rawValue) / 10.0;
                channels[idxC].retVal      := 16#0000;

            2: (* ---- Climatic‑temperature conversion ---- *)
                channels[idxC].outputValue := INT_TO_REAL(rawValue) / 100.0;
                channels[idxC].retVal      := 16#0000;

            ELSE
                (* Unknown measuring mode *)
                channels[idxC].retVal      := 16#8001;  (* Invalid mode *)
                channels[idxC].outputValue := 0.0;
        END_CASE

    END_FOR
END_FUNCTION_BLOCK

(* ---- public-medium-02.candidate_02.st ---- *)
(*--------------------------------------------------------------
  Type definition for a single analog channel.
--------------------------------------------------------------*)
TYPE ST_AnalogChannel
STRUCT
    enable        : BOOL;      (* Channel conversion enable *)
    hiLIM         : REAL;      (* Upper engineering-unit limit *)
    loLIM         : REAL;      (* Lower engineering-unit limit *)
    bipolar       : BOOL;      (* FALSE → unipolar, TRUE → bipolar *)
    measuringMode : INT;       (* 0 = linear, 1 = std temp, 2 = climatic *)
    retVal        : WORD;      (* Per-channel status code (output) *)
    outputValue   : REAL;      (* Converted engineering value (output) *)
END_STRUCT
END_TYPE

(*--------------------------------------------------------------
  Function block: FB_AnalogBatchProcessing
  Processes up to *count* analog channels.
--------------------------------------------------------------*)
FUNCTION_BLOCK FB_AnalogBatchProcessing
VAR_INPUT
    count : DINT;                      (* Number of channels to process *)
END_VAR
VAR_IN_OUT
    analogValues : ARRAY[*] OF INT;    (* Raw analog values (read-only) *)
    channels     : ARRAY[*] OF ST_AnalogChannel; (* Channel settings & results *)
END_VAR
VAR
    i          : DINT;
    rawValue   : INT;
    rawMin     : REAL;
    rawMax     : REAL;
    scale      : REAL;
    ch         : ST_AnalogChannel;
END_VAR

    FOR i := 0 TO count - 1 DO
        rawValue := analogValues[LOWER_BOUND(analogValues, 1) + i];
        ch := channels[LOWER_BOUND(channels, 1) + i];

        IF NOT ch.enable THEN
            channels[LOWER_BOUND(channels, 1) + i].retVal      := 16#0000;
            channels[LOWER_BOUND(channels, 1) + i].outputValue := 0.0;
        ELSE
            CASE ch.measuringMode OF
                0: (* ---- Non-temperature linear scaling ---- *)
                    IF ch.hiLIM <= ch.loLIM THEN
                        channels[LOWER_BOUND(channels, 1) + i].retVal      := 16#8002;
                        channels[LOWER_BOUND(channels, 1) + i].outputValue := 0.0;
                    ELSE
                        IF ch.bipolar THEN
                            rawMin := -27648.0;
                            rawMax :=  27648.0;
                        ELSE
                            rawMin := 0.0;
                            rawMax := 27648.0;
                        END_IF
                        scale := (ch.hiLIM - ch.loLIM) / (rawMax - rawMin);
                        channels[LOWER_BOUND(channels, 1) + i].outputValue := ch.loLIM
                                     + (INT_TO_REAL(rawValue) - rawMin) * scale;
                        channels[LOWER_BOUND(channels, 1) + i].retVal := 16#0000;
                    END_IF

                1: (* ---- Standard-temperature conversion ---- *)
                    channels[LOWER_BOUND(channels, 1) + i].outputValue := INT_TO_REAL(rawValue) / 10.0;
                    channels[LOWER_BOUND(channels, 1) + i].retVal      := 16#0000;

                2: (* ---- Climatic-temperature conversion ---- *)
                    channels[LOWER_BOUND(channels, 1) + i].outputValue := INT_TO_REAL(rawValue) / 100.0;
                    channels[LOWER_BOUND(channels, 1) + i].retVal      := 16#0000;

                ELSE
                    channels[LOWER_BOUND(channels, 1) + i].retVal      := 16#8001;
                    channels[LOWER_BOUND(channels, 1) + i].outputValue := 0.0;
            END_CASE
        END_IF
    END_FOR
END_FUNCTION_BLOCK

(* ---- public-medium-03.candidate_01.st ---- *)
FUNCTION_BLOCK FB_MovingAverage
VAR_INPUT
    cyclicExecution  : BOOL;  // When TRUE, periodic reading is performed
    trigger          : BOOL;  // External trigger signal, reads value upon each rising edge
    value            : LREAL; // Newly read data value
    windowSize       : INT;   // Window size for moving average (1-100)
    reset            : BOOL;  // Reset signal, resets the moving average calculation when TRUE
END_VAR

VAR_OUTPUT
    average          : LREAL; // The moving average result
    windowSizeReached: BOOL;  // FALSE: Maximum window width not yet reached
                              // TRUE: Maximum window width has been reached
    error            : BOOL;  // FALSE: No error occurred, TRUE: An error occurred
    status           : WORD;  // Status code
END_VAR

VAR
    dataBuffer       : ARRAY[1..100] OF LREAL; // Circular buffer for data values
    sum              : LREAL;                   // Sum of values in current window
    validSampleCount : INT;                     // Number of valid samples in buffer
    prevTrigger      : BOOL;                    // Previous trigger state for edge detection
END_VAR

// ============================================================================
// Reset Handling
// ============================================================================
IF reset THEN
    sum              := 0.0;
    validSampleCount := 0;
    average          := 0.0;
    windowSizeReached := FALSE;
    error            := FALSE;
    status           := 16#0000;
    prevTrigger      := FALSE;
    RETURN;
END_IF

// ============================================================================
// Window Size Validation
// ============================================================================
IF windowSize < 1 OR windowSize > 100 THEN
    error  := TRUE;
    status := 16#8200;  // Window length setting error
    RETURN;
END_IF

// Clear error on successful validation
error  := FALSE;
status := 16#0000;     // Execution successful

// ============================================================================
// Process New Value
// Condition: cyclicExecution is TRUE OR trigger has a rising edge
// ============================================================================
IF cyclicExecution OR (trigger AND NOT prevTrigger) THEN
    // When buffer is full, remove the oldest value from sum
    IF validSampleCount >= windowSize THEN
        sum := sum - dataBuffer[1];

        // Shift buffer elements left (simple shifting approach)
        FOR i := 1 TO windowSize - 1 DO
            dataBuffer[i] := dataBuffer[i + 1];
        END_FOR
    END_IF

    // Add new value to buffer
    dataBuffer[validSampleCount + 1] := value;
    sum := sum + value;

    // Update sample count (max is windowSize)
    IF validSampleCount < windowSize THEN
        validSampleCount := validSampleCount + 1;
    END_IF

    // Calculate average
    average := sum / INT_TO_LREAL(validSampleCount);

    // Check if window has been filled to maximum size
    windowSizeReached := (validSampleCount = windowSize);
END_IF

// ============================================================================
// Update Trigger State for Rising Edge Detection
// ============================================================================
prevTrigger := trigger;

END_FUNCTION_BLOCK

(* ---- public-medium-03.candidate_02.st ---- *)
FUNCTION_BLOCK FB_MovingAverage
VAR_INPUT
    cyclicExecution  : BOOL;  // When TRUE, periodic reading is performed
    trigger          : BOOL;  // External trigger signal, reads value upon each rising edge
    value            : LREAL; // Newly read data value
    windowSize       : INT;   // Window size for moving average (1-100)
    reset            : BOOL;  // Reset signal, resets the moving average calculation when TRUE
END_VAR

VAR_OUTPUT
    average          : LREAL; // The moving average result
    windowSizeReached: BOOL;  // FALSE: Maximum window width not yet reached
                              // TRUE: Maximum window width has been reached
    error            : BOOL;  // FALSE: No error occurred, TRUE: An error occurred
    status           : WORD;  // Status code
END_VAR

VAR
    dataBuffer       : ARRAY[1..100] OF LREAL; // Circular buffer for data values
    sum              : LREAL;                   // Sum of values in current window
    validSampleCount : INT;                     // Number of valid samples in buffer
    prevTrigger      : BOOL;                    // Previous trigger state for edge detection
    i                : INT;                     // Loop counter
END_VAR

// ============================================================================
// Reset Handling
// ============================================================================
IF reset THEN
    sum              := 0.0;
    validSampleCount := 0;
    average          := 0.0;
    windowSizeReached := FALSE;
    error            := FALSE;
    status           := 16#0000;
    prevTrigger      := FALSE;
    RETURN;
END_IF

// ============================================================================
// Window Size Validation
// ============================================================================
IF windowSize < 1 OR windowSize > 100 THEN
    error  := TRUE;
    status := 16#8200;  // Window length setting error
    RETURN;
END_IF

// Clear error on successful validation
error  := FALSE;
status := 16#0000;     // Execution successful

// ============================================================================
// Process New Value
// Condition: cyclicExecution is TRUE OR trigger has a rising edge
// ============================================================================
IF cyclicExecution OR (trigger AND NOT prevTrigger) THEN
    // When buffer is full, remove the oldest value from sum
    IF validSampleCount >= windowSize THEN
        sum := sum - dataBuffer[1];

        // Shift buffer elements left
        FOR i := 1 TO windowSize - 1 DO
            dataBuffer[i] := dataBuffer[i + 1];
        END_FOR
    END_IF

    // Add new value to buffer
    dataBuffer[validSampleCount + 1] := value;
    sum := sum + value;

    // Update sample count (max is windowSize)
    IF validSampleCount < windowSize THEN
        validSampleCount := validSampleCount + 1;
    END_IF

    // Calculate average
    average := sum / INT_TO_LREAL(validSampleCount);

    // Check if window has been filled to maximum size
    windowSizeReached := (validSampleCount = windowSize);
END_IF

// ============================================================================
// Update Trigger State for Rising Edge Detection
// ============================================================================
prevTrigger := trigger;

END_FUNCTION_BLOCK

(* ---- public-medium-04.candidate_01.st ---- *)
(*====================================================================*)
(*  FUNCTION_BLOCK FB_TemperatureControl                              *)
(*  Implements a temperature‑control loop with over‑heat protection   *)
(*  and sensor‑fault detection.                                       *)
(*                                                                    *)
(*  Inputs:                                                           *)
(*    TemperatureSensorInput  – REAL  – actual temperature (°C)       *)
(*    SetTemperature          – REAL  – desired temperature (°C)      *)
(*                                                                    *)
(*  Outputs:                                                          *)
(*    CurrentTemperature      – REAL  – display of current temperature*)
(*    SetTempDisplay          – REAL  – display of set temperature    *)
(*    HeaterStatus            – BOOL  – heater ON/OFF status          *)
(*    OverheatProtection      – BOOL  – over‑heat protection active   *)
(*    HeaterOutput            – BOOL  – heater control output         *)
(*====================================================================*)

FUNCTION_BLOCK FB_TemperatureControl

VAR_INPUT
    TemperatureSensorInput : REAL;   (* Actual temperature from sensor *)
    SetTemperature         : REAL;   (* Desired temperature set point  *)
END_VAR

VAR_OUTPUT
    CurrentTemperature : REAL;       (* Display of current temperature *)
    SetTempDisplay     : REAL;       (* Display of set temperature      *)
    HeaterStatus       : BOOL;       (* Heater ON/OFF status            *)
    OverheatProtection : BOOL;       (* Over‑heat protection flag       *)
    HeaterOutput       : BOOL;       (* Heater control output           *)
END_VAR

VAR
    (* Internal control signals *)
    HeatingRequested   : BOOL;       (* TRUE when heating is required   *)
    SensorFault        : BOOL;       (* TRUE when sensor reading is out‑of‑range *)

    (* Timer instances *)
    OverheatTimer      : TON;        (* Counts ON‑time of the heater     *)
    OverheatWaitTimer  : TON;        (* Counts the 3 s wait after over‑heat *)
END_VAR

(*------------------------------------------------------------------*)
(* 1. Sensor‑fault detection (0 °C … 100 °C is the valid range)      *)
(*------------------------------------------------------------------*)
SensorFault := (TemperatureSensorInput < 0.0) OR (TemperatureSensorInput > 100.0);

(*------------------------------------------------------------------*)
(* 2. Determine if heating is required (based on temperature)        *)
(*------------------------------------------------------------------*)
IF SensorFault THEN
    HeatingRequested := FALSE;                 (* Fault → no heating *)
ELSE
    IF TemperatureSensorInput < SetTemperature THEN
        HeatingRequested := TRUE;              (* Below set point → heat *)
    ELSE
        HeatingRequested := FALSE;             (* At or above set point   *)
    END_IF
END_IF

(*------------------------------------------------------------------*)
(* 3. Over‑heat detection timer (5 s continuous heater ON)           *)
(*------------------------------------------------------------------*)
OverheatTimer(IN := HeaterOutput, PT := T#5s);

(* If the timer elapses while protection is not yet active,          *)
(* raise the protection flag and force the heater OFF immediately.   *)
IF OverheatTimer.Q AND NOT OverheatProtection THEN
    OverheatProtection := TRUE;
    HeaterOutput       := FALSE;                (* Ensure heater is off   *)
END_IF

(*------------------------------------------------------------------*)
(* 4. Over‑heat wait timer (3 s must elapse before protection can be cleared) *)
(*------------------------------------------------------------------*)
OverheatWaitTimer(IN := OverheatProtection, PT := T#3s);

(* After the mandatory 3 s wait, clear the protection flag.          *)
IF OverheatWaitTimer.Q THEN
    OverheatProtection := FALSE;
END_IF

(*------------------------------------------------------------------*)
(* 5. Final heater command – allowed only when heating is requested  *)
(*    and over‑heat protection is NOT active.                        *)
(*------------------------------------------------------------------*)
HeaterOutput := HeatingRequested AND NOT OverheatProtection;

(*------------------------------------------------------------------*)
(* 6. Status outputs                                                *)
(*------------------------------------------------------------------*)
CurrentTemperature := TemperatureSensorInput;   (* Display current temp *)
SetTempDisplay     := SetTemperature;           (* Display set temp     *)
HeaterStatus       := HeaterOutput;             (* Heater ON/OFF status *)

END_FUNCTION_BLOCK
(*====================================================================*)

(* ---- public-medium-05.candidate_02.st ---- *)
FUNCTION_BLOCK ProductionLineControl
VAR_INPUT
    Mode            : BOOL;   // 0=manual mode, 1=automatic mode
    ForwardButton   : BOOL;   // Forward rotation button
    ReverseButton   : BOOL;   // Reverse rotation button
    SensorA         : BOOL;   // Sensor A
    SensorB         : BOOL;   // Sensor B
    SensorC         : BOOL;   // Sensor C
    ButtonA         : BOOL;   // Button A
    ButtonB         : BOOL;   // Button B
    ButtonC         : BOOL;   // Button C
END_VAR

VAR_OUTPUT
    MotorForward    : BOOL;   // Motor forward rotation output
    MotorReverse    : BOOL;   // Motor reverse rotation output
    CompletionLight : BOOL;   // Indicator light for product processing completion
END_VAR

VAR
    State           : INT := 0;  // 0=WAIT_A, 1=WAIT_A_PRESSED, 2=MOVING_AB, 3=WAIT_B_PRESSED, 4=MOVING_BC, 5=WAIT_C_PRESSED, 6=COMPLETE
    SensorA_Prev    : BOOL := FALSE;
    SensorB_Prev    : BOOL := FALSE;
    SensorC_Prev    : BOOL := FALSE;
END_VAR

// Edge detection for sensors
VAR
    SensorA_Edge    : BOOL;
    SensorB_Edge    : BOOL;
    SensorC_Edge    : BOOL;
END_VAR

SensorA_Edge := SensorA AND NOT SensorA_Prev;
SensorB_Edge := SensorB AND NOT SensorB_Prev;
SensorC_Edge := SensorC AND NOT SensorC_Prev;

// Store previous sensor states for edge detection
SensorA_Prev := SensorA;
SensorB_Prev := SensorB;
SensorC_Prev := SensorC;

// Manual Mode (Mode = 0)
IF Mode = FALSE THEN
    // Reset state to initial when switching to manual mode
    State := 0;

    // Forward and reverse rotation with interlock
    MotorForward := ForwardButton AND NOT ReverseButton;
    MotorReverse := ReverseButton AND NOT ForwardButton;

    // Completion light is off in manual mode
    CompletionLight := FALSE;

// Automatic Mode (Mode = 1)
ELSE
    // State machine logic
    CASE State OF
        // State 0: Waiting for product at Workstation A
        0:  // WAIT_A
            MotorForward := FALSE;
            MotorReverse := FALSE;

            // Detect product arrival at A
            IF SensorA_Edge THEN
                State := 1;
            END_IF

        // State 1: Product at A, waiting for operator to press ButtonA
        1:  // WAIT_A_PRESSED
            MotorForward := FALSE;
            MotorReverse := FALSE;

            // Operator presses ButtonA to signal processing complete
            IF ButtonA THEN
                State := 2;
            END_IF

            // Safety: If product leaves A unexpectedly, return to WAIT_A
            IF NOT SensorA THEN
                State := 0;
            END_IF

        // State 2: Motor moving product from A to B
        2:  // MOVING_AB
            MotorForward := TRUE;
            MotorReverse := FALSE;

            // Product arrives at B
            IF SensorB THEN
                State := 3;
            END_IF

        // State 3: Product at B, waiting for operator to press ButtonB
        3:  // WAIT_B_PRESSED
            MotorForward := FALSE;
            MotorReverse := FALSE;

            // Operator presses ButtonB to signal processing complete
            IF ButtonB THEN
                State := 4;
            END_IF

            // Safety: If product leaves B unexpectedly, return to WAIT_A
            IF NOT SensorB THEN
                State := 0;
            END_IF

        // State 4: Motor moving product from B to C
        4:  // MOVING_BC
            MotorForward := TRUE;
            MotorReverse := FALSE;

            // Product arrives at C
            IF SensorC THEN
                State := 5;
            END_IF

        // State 5: Product at C, waiting for operator to press ButtonC
        5:  // WAIT_C_PRESSED
            MotorForward := FALSE;
            MotorReverse := FALSE;

            // Operator presses ButtonC to signal processing complete
            IF ButtonC THEN
                State := 6;
            END_IF

            // Safety: If product leaves C unexpectedly, return to WAIT_A
            IF NOT SensorC THEN
                State := 0;
            END_IF

        // State 6: Product processing complete
        6:  // COMPLETE
            MotorForward := FALSE;
            MotorReverse := FALSE;

            // When product is taken away (SensorC no longer detects product)
            IF NOT SensorC THEN
                State := 0;
            END_IF

    END_CASE;

    // Set CompletionLight based on current state
    CompletionLight := (State = 6);

END_IF;

END_FUNCTION_BLOCK

(* ---- public-medium-07.candidate_02.st ---- *)
(* -------------------------------------------------------------
   Office HVAC Multi‑mode Energy‑Saving Control
   -------------------------------------------------------------
   Inputs
     OCCUPANCY_DETECTED   – TRUE when occupancy is detected
     ENERGY_SAVING_MODE   – TRUE → energy‑saving, FALSE → standard
     HVAC_MODE_SELECTOR   – 0 = Auto, 1 = Comfort, 2 = Economy, 3 = Night
   Outputs
     SUPPLY_FAN_RUN       – Supply‑fan run enable (BOOL)
     TEMP_SETPOINT_ADJUST – Temperature‑setpoint adjustment in °C (INT)
   -------------------------------------------------------------
   Behaviour
     • 30 s on‑delay for the fan when occupied and NOT in Night mode.
       The fan is stopped immediately and the timer is reset when
       occupancy is lost or Night mode is entered.
     • Temperature‑setpoint adjustment follows the table:
       Mode   | Occupied | Unoccupied (standard) | Unoccupied (energy‑saving)
       -------|----------|-----------------------|----------------------------
       Auto   |   0 °C   |        +2 °C          |            +3 °C
       Comfort|   0 °C   |        +1 °C          |            +1 °C
       Economy|   0 °C   |        +4 °C          |            +4 °C
       Night  |   +4 °C  |        +4 °C          |            +4 °C
       (Energy‑saving flag influences only Auto mode.)
     • Outputs are initialised to OFF / 0 at power‑up and are updated
       every scan from the current inputs.
   ------------------------------------------------------------- *)

FUNCTION_BLOCK HVAC_Control
   VAR_INPUT
      OCCUPANCY_DETECTED   : BOOL;
      ENERGY_SAVING_MODE   : BOOL;
      HVAC_MODE_SELECTOR   : INT;
   END_VAR

   VAR_OUTPUT
      SUPPLY_FAN_RUN       : BOOL := FALSE;
      TEMP_SETPOINT_ADJUST : INT  := 0;
   END_VAR

   VAR
      FanTimer      : TON;
      FanStartCond  : BOOL;
   END_VAR

   (* ---------------------------------------------------------
      Fan start condition: occupied AND NOT Night mode
      --------------------------------------------------------- *)
   FanStartCond := OCCUPANCY_DETECTED AND (HVAC_MODE_SELECTOR <> 3);

   (* ---------------------------------------------------------
      30‑second ON‑delay timer
      The timer resets automatically when FanStartCond becomes FALSE,
      fulfilling the “reset timing if occupancy is lost or Night mode
      is selected” requirement.
      --------------------------------------------------------- *)
   FanTimer(IN := FanStartCond, PT := T#30s);
   SUPPLY_FAN_RUN := FanTimer.Q;

   (* ---------------------------------------------------------
      Temperature‑setpoint adjustment according to mode,
      occupancy and energy‑saving selection.
      --------------------------------------------------------- *)
   CASE HVAC_MODE_SELECTOR OF
      0 : (* Auto *)
         IF OCCUPANCY_DETECTED THEN
            TEMP_SETPOINT_ADJUST := 0;
         ELSE
            IF ENERGY_SAVING_MODE THEN
               TEMP_SETPOINT_ADJUST := 3;
            ELSE
               TEMP_SETPOINT_ADJUST := 2;
            END_IF;
         END_IF;

      1 : (* Comfort *)
         IF OCCUPANCY_DETECTED THEN
            TEMP_SETPOINT_ADJUST := 0;
         ELSE
            TEMP_SETPOINT_ADJUST := 1;
         END_IF;

      2 : (* Economy *)
         IF OCCUPANCY_DETECTED THEN
            TEMP_SETPOINT_ADJUST := 0;
         ELSE
            TEMP_SETPOINT_ADJUST := 4;
         END_IF;

      3 : (* Night *)
         TEMP_SETPOINT_ADJUST := 4;

   END_CASE;

END_FUNCTION_BLOCK

(* ---- public-medium-08.candidate_01.st ---- *)
FUNCTION_BLOCK FB_ParseIPv4
VAR_INPUT
    ipText : STRING(254);
END_VAR
VAR_OUTPUT
    ipValue : UDINT;
END_VAR
VAR
    i           : INT;
    length      : INT;
    segmentIdx  : INT;
    segValue    : UDINT;
    isValid     : BOOL;
    ch          : BYTE;
    digit       : BYTE;
    segments    : ARRAY[0..3] OF UDINT;
END_VAR

// Initialize output to invalid state
ipValue := 0;

// Reset parsing state
isValid    := TRUE;
segmentIdx := 0;
segValue   := 0;
length     := LEN(ipText);

// Empty input check
IF length = 0 THEN
    RETURN;
END_IF

// Parse through each character
FOR i := 1 TO length DO
    ch := BYTE_TO_INT(CHAR_TO_BYTE(MID(ipText, 1, i)));

    // Digit: 0-9 ASCII range 48-57
    IF ch >= 48 AND ch <= 57 THEN
        digit := ch - 48;

        // Check for overflow before multiplying
        // Max valid segment is 255
        // If current value > 25, multiplying by 10 would exceed 255
        // If current value = 25, digit > 5 would exceed 255
        IF segValue > 25 OR (segValue = 25 AND digit > 5) THEN
            isValid := FALSE;
            EXIT;
        END_IF;

        segValue := segValue * 10 + digit;

    // Period: segment delimiter
    ELSIF ch = 46 THEN
        IF segmentIdx > 3 THEN
            isValid := FALSE;
            EXIT;
        END_IF;

        segments[segmentIdx] := segValue;
        segmentIdx := segmentIdx + 1;
        segValue   := 0;

    // Any other character is invalid
    ELSE
        isValid := FALSE;
        EXIT;
    END_IF
END_FOR

// Process final segment
IF isValid THEN
    IF segmentIdx > 3 THEN
        isValid := FALSE;
    ELSE
        segments[segmentIdx] := segValue;
        segmentIdx := segmentIdx + 1;
    END_IF
END_IF

// Validate exactly 4 segments
IF isValid AND segmentIdx <> 4 THEN
    isValid := FALSE;
END_IF

// Assemble result in network byte order (MSB first)
// ipValue[31:24] = segments[0]
// ipValue[23:16] = segments[1]
// ipValue[15:8]  = segments[2]
// ipValue[7:0]   = segments[3]
IF isValid THEN
    ipValue := SHL(segments[0], 24) OR SHL(segments[1], 16)
             OR SHL(segments[2], 8)  OR segments[3];
ELSE
    ipValue := 0;
END_IF

END_FUNCTION_BLOCK

(* ---- public-medium-08.candidate_02.st ---- *)
FUNCTION_BLOCK FB_ParseIPv4
VAR_INPUT
    ipText : STRING(254);
END_VAR
VAR_OUTPUT
    ipValue : UDINT;
END_VAR
VAR
    i           : INT;
    length      : INT;
    segmentIdx  : INT;
    segValue    : UDINT;
    isValid     : BOOL;
    curChar     : STRING(1);
    segments    : ARRAY[0..3] OF UDINT;
END_VAR

// Initialize output to invalid state
ipValue := 0;
isValid := TRUE;
segmentIdx := 0;
segValue := 0;
length := LEN(ipText);

// Empty input check
IF length = 0 THEN
    RETURN;
END_IF

// Parse through each character
FOR i := 1 TO length DO
    curChar := MID(ipText, 1, i);

    // Digit check: compare STRING(1) to character literals
    IF curChar = '0' OR curChar = '1' OR curChar = '2' OR
       curChar = '3' OR curChar = '4' OR curChar = '5' OR
       curChar = '6' OR curChar = '7' OR curChar = '8' OR
       curChar = '9' THEN

        // Check for overflow before accumulating
        IF segValue > 25 OR (segValue = 25 AND curChar > '5') THEN
            isValid := FALSE;
            EXIT;
        END_IF;

        // Accumulate digit value (convert char to numeric)
        IF curChar = '0' THEN segValue := segValue * 10 + 0;
        ELSIF curChar = '1' THEN segValue := segValue * 10 + 1;
        ELSIF curChar = '2' THEN segValue := segValue * 10 + 2;
        ELSIF curChar = '3' THEN segValue := segValue * 10 + 3;
        ELSIF curChar = '4' THEN segValue := segValue * 10 + 4;
        ELSIF curChar = '5' THEN segValue := segValue * 10 + 5;
        ELSIF curChar = '6' THEN segValue := segValue * 10 + 6;
        ELSIF curChar = '7' THEN segValue := segValue * 10 + 7;
        ELSIF curChar = '8' THEN segValue := segValue * 10 + 8;
        ELSIF curChar = '9' THEN segValue := segValue * 10 + 9;
        END_IF

    // Period: segment delimiter
    ELSIF curChar = '.' THEN
        IF segmentIdx >= 4 THEN
            isValid := FALSE;
            EXIT;
        END_IF;

        segments[segmentIdx] := segValue;
        segmentIdx := segmentIdx + 1;
        segValue := 0;

    // Any other character is invalid
    ELSE
        isValid := FALSE;
        EXIT;
    END_IF
END_FOR

// Process final segment
IF isValid THEN
    IF segmentIdx >= 4 THEN
        isValid := FALSE;
    ELSE
        segments[segmentIdx] := segValue;
        segmentIdx := segmentIdx + 1;
    END_IF
END_IF

// Validate exactly 4 segments
IF isValid AND segmentIdx <> 4 THEN
    isValid := FALSE;
END_IF

// Assemble result in network byte order (MSB first)
IF isValid THEN
    ipValue := SHL(segments[0], 24) OR SHL(segments[1], 16)
             OR SHL(segments[2], 8)  OR segments[3];
ELSE
    ipValue := 0;
END_IF

END_FUNCTION_BLOCK

(* ---- self-easy-01.candidate_01.st ---- *)
FUNCTION_BLOCK FB
VAR_INPUT
    enable     : BOOL;               (* TRUE → update average, FALSE → keep previous *)
    values     : ARRAY[1..8] OF INT; (* sampled raw values (1..8 stations) *)
    count      : INT;                (* number of valid samples this cycle (0..8) *)
    avgEnable  : BOOL;               (* averaging enable – when FALSE keep previous *)
END_VAR
VAR_OUTPUT
    avgOut     : REAL;               (* average output *)
END_VAR
VAR
    lastAvg        : REAL := 0.0;    (* stores the previous average for retention *)
    sum            : DINT;           (* wider type to avoid overflow while summing *)
    i              : INT;
    effectiveCount : INT;            (* count limited to the array size 8 *)
END_VAR

(* ---------------------------------------------------------------
   Compute the arithmetic mean of the first ‘effectiveCount’
   samples when:
      • enable      = TRUE
      • avgEnable   = TRUE
      • count       > 0
   In all other situations the output is held at its previous
   value (lastAvg).  No division‑by‑zero can occur because the
   guard “count > 0” is tested before the division.
   --------------------------------------------------------------- *)
IF enable AND avgEnable AND count > 0 THEN
    (* clip count to the available array length *)
    effectiveCount := count;
    IF effectiveCount > 8 THEN
        effectiveCount := 8;
    END_IF;

    (* sum the first ‘effectiveCount’ values using DINT *)
    sum := 0;
    FOR i := 1 TO effectiveCount DO
        sum := sum + values[i];
    END_FOR;

    (* compute the average as REAL (no rounding) *)
    avgOut    := DINT_TO_REAL(sum) / DINT_TO_REAL(effectiveCount);
    lastAvg   := avgOut;          (* remember for cycles where we keep the value *)
ELSE
    (* keep the previous average *)
    avgOut    := lastAvg;
END_IF;

END_FUNCTION_BLOCK

(* ---- self-easy-02.candidate_01.st ---- *)
FUNCTION_BLOCK FB
VAR_INPUT
    tankLevel   : REAL;
    outletFlow  : REAL;
    inletPermit : BOOL;
    resetBtn    : BOOL;
END_VAR

VAR_OUTPUT
    pumpRun         : BOOL;
    alarmHigh       : BOOL;
    alarmLow        : BOOL;
    outletValveOpen : BOOL;
END_VAR

VAR
    prevResetBtn  : BOOL := FALSE;
    prevAlarmHigh : BOOL := FALSE;
    prevAlarmLow  : BOOL := FALSE;

    risingReset : BOOL;
    highHazard  : BOOL;
    lowHazard   : BOOL;
END_VAR

(* 检測複位按鍵上升沿 *)
risingReset := resetBtn AND NOT prevResetBtn;

(* 危險條件 *)
highHazard := (tankLevel >= 85.0);
lowHazard  := (tankLevel <= 15.0);

(* 報警鎖存：危險條件成立時立即置位，否則跟隨上一拍狀態（若未出現復位上升沿） *)
alarmHigh := highHazard OR (prevAlarmHigh AND NOT risingReset);
alarmLow  := lowHazard  OR (prevAlarmLow  AND NOT risingReset);

(* 輸出 *)
pumpRun         := inletPermit AND NOT alarmHigh AND NOT alarmLow;
outletValveOpen := NOT alarmLow;

(* 為下一掃描保存狀態 *)
prevResetBtn  := resetBtn;
prevAlarmHigh := alarmHigh;
prevAlarmLow  := alarmLow;

END_FUNCTION_BLOCK

(* ---- self-hard-01.candidate_01.st ---- *)
FUNCTION_BLOCK FB
VAR_INPUT
    flowLow : BOOL;
    ackBtn : BOOL;
    sensorOK : BOOL;
END_VAR
VAR_OUTPUT
    alarmActive : BOOL;
    alarmAcked : BOOL;
    highHigh : BOOL;
END_VAR
VAR
    prev_flowLow : BOOL := FALSE;
    prev_ackBtn : BOOL := FALSE;
END_VAR

// 高优先级报警：传感器断线时置位
highHigh := NOT sensorOK;

// 检测确认按钮上升沿
VAR rising : BOOL;
rising := ackBtn AND NOT prev_ackBtn;

// 计算新的报警状态（基于形式化性质）
VAR newAlarmActive : BOOL;
VAR newAlarmAcked : BOOL;

newAlarmActive := flowLow OR (alarmActive AND NOT rising AND NOT (prev_flowLow AND alarmAcked));

newAlarmAcked := newAlarmActive AND (NOT flowLow OR rising OR (prev_flowLow AND alarmActive AND alarmAcked));

alarmActive := newAlarmActive;
alarmAcked := newAlarmAcked;

// 更新历史变量
prev_flowLow := flowLow;
prev_ackBtn := ackBtn;

END_FUNCTION_BLOCK

(* ---- self-hard-01.candidate_02.st ---- *)
FUNCTION_BLOCK FB
VAR_INPUT
    flowLow  : BOOL;
    ackBtn   : BOOL;
    sensorOK : BOOL;
END_VAR
VAR_OUTPUT
    alarmActive : BOOL;
    alarmAcked  : BOOL;
    highHigh    : BOOL;
END_VAR
VAR
    prevFlowLow : BOOL := FALSE;
    prevAckBtn  : BOOL := FALSE;
    risingEdge  : BOOL;
END_VAR

// S5: highHigh 与传感器状态双向一致
highHigh := NOT sensorOK;

// S4: 检测确认按钮上升沿
risingEdge := ackBtn AND NOT prevAckBtn;

// S1/S2/S6: 报警激活逻辑
// flowLow出现则激活；已激活且未确认时不消失；条件消失后仅确认沿清除
alarmActive := flowLow OR (alarmActive AND NOT risingEdge AND NOT (prevFlowLow AND alarmAcked));

// S4/S7: 报警已确认逻辑
// 条件消失后自动置位；确认沿出现且条件仍在时置位；保持记忆状态
alarmAcked := alarmActive AND (NOT flowLow OR risingEdge OR (prevFlowLow AND alarmAcked));

// 更新历史变量
prevFlowLow := flowLow;
prevAckBtn  := ackBtn;

END_FUNCTION_BLOCK

(* ---- self-hard-02.candidate_01.st ---- *)
FUNCTION_BLOCK FB
VAR_INPUT
    startBtn    : BOOL;
    abortBtn    : BOOL;
    setpoint    : REAL;
    pv          : REAL;
    maxDuration : INT;
END_VAR
VAR_OUTPUT
    elapsed : INT;
    phase   : INT;
    timeout : BOOL;
END_VAR
VAR
    prevStartBtn : BOOL := FALSE;
    prevPhase    : INT  := 0;
    prevElapsed  : INT  := 0;
    prevTimeout  : BOOL := FALSE;
END_VAR

(* temporary variable for rising edge detection *)
VAR
    risingStart : BOOL;
END_VAR

(* detect rising edge of start button *)
risingStart := startBtn AND NOT prevStartBtn;

(* abort has the highest priority *)
IF abortBtn THEN
    phase   := 9;
    elapsed := prevElapsed;
    timeout := prevTimeout;
    (* the start‑button rising edge in this scan is ignored *)
ELSE
    (* new batch start on rising edge of start button *)
    IF risingStart THEN
        phase   := 1;
        elapsed := 0;
        timeout := FALSE;
    ELSE
        (* no abort, no new start: update based on previous state *)
        IF (prevPhase = 1) OR (prevPhase = 2) THEN
            (* running phase – increment scan counter *)
            elapsed := prevElapsed + 1;

            (* check for timeout *)
            IF elapsed >= maxDuration THEN
                timeout := TRUE;
                phase   := 3;                (* completed due to timeout *)
            ELSE
                (* no timeout – decide heating or holding according to temperature *)
                IF prevPhase = 1 THEN
                    IF pv >= setpoint THEN
                        phase := 2;          (* temperature reached → hold *)
                    ELSE
                        phase := 1;          (* still heating *)
                    END_IF;
                ELSE                           (* prevPhase = 2 *)
                    phase := 2;              (* remain in holding *)
                END_IF;
                timeout := prevTimeout;       (* should be FALSE *)
            END_IF;
        ELSE
            (* previous scan was not a running phase – keep state unchanged *)
            phase   := prevPhase;
            elapsed := prevElapsed;
            timeout := prevTimeout;
        END_IF;
    END_IF;
END_IF;

(* update memory for the next scan *)
prevStartBtn := startBtn;
prevPhase    := phase;
prevElapsed  := elapsed;
prevTimeout  := timeout;

END_FUNCTION_BLOCK

(* ---- self-hard-03.candidate_01.st ---- *)
FUNCTION_BLOCK FB
VAR_INPUT
    pushEn  : BOOL;          // 入队指令（上升沿有效）
    pushItem: INT;           // 入队物料号
    popEn   : BOOL;          // 出队指令（上升沿有效）
END_VAR
VAR_INOUT
    fifo : ARRAY[1..8] OF INT; // 队列缓冲区，下标 1 为最老元素
END_VAR
VAR_OUTPUT
    count : INT;             // 当前队列元素个数 0..8
    full  : BOOL;            // 队列满
    empty : BOOL;            // 队列空
    head  : INT;             // 队首元素（空时保持 0）
END_VAR
VAR
    prevPush : BOOL := FALSE; // 上一周期 pushEn 的状态
    prevPop  : BOOL := FALSE; // 上一周期 popEn 的状态
    i        : INT;          // 循环计数器
END_VAR

    // ------------------------------------------------------------
    // 1. 出队：popEn 上升沿先执行（仅在队列非空时有效）
    // ------------------------------------------------------------
    IF popEn AND NOT prevPop THEN
        IF count > 0 THEN
            // 将所有有效元素左移一位，实现移除 fifo[1]
            FOR i := 1 TO count - 1 DO
                fifo[i] := fifo[i + 1];
            END_FOR
            // 将被腾出的最后一个位置清零（可选，满足“紧凑”要求）
            fifo[count] := 0;
            count := count - 1;
        END_IF
    END_IF

    // ------------------------------------------------------------
    // 2. 入队：pushEn 上升沿随后执行（仅在队列未满时有效）
    // ------------------------------------------------------------
    IF pushEn AND NOT prevPush THEN
        IF count < 8 THEN
            count := count + 1;
            fifo[count] := pushItem;   // 新元素追加到逻辑队尾
        END_IF
    END_IF

    // ------------------------------------------------------------
    // 3. 输出信号
    // ------------------------------------------------------------
    full  := (count = 8);
    empty := (count = 0);
    head  := 0;
    IF NOT empty THEN
        head := fifo[1];
    END_IF

    // ------------------------------------------------------------
    // 4. 更新历史状态，供下一周期边沿检测使用
    // ------------------------------------------------------------
    prevPush := pushEn;
    prevPop  := popEn;
END_FUNCTION_BLOCK

(* ---- self-hard-03.candidate_02.st ---- *)
FUNCTION_BLOCK FB
VAR_INPUT
    pushEn  : BOOL;
    pushItem: INT;
    popEn   : BOOL;
END_VAR
VAR_IN_OUT
    fifo : ARRAY[1..8] OF INT;
END_VAR
VAR_OUTPUT
    count : INT;
    full  : BOOL;
    empty : BOOL;
    head  : INT;
END_VAR
VAR
    prevPush : BOOL;
    prevPop  : BOOL;
    i        : INT;
END_VAR

    // pop rising edge: remove first element if not empty
    IF popEn AND NOT prevPop THEN
        IF count > 0 THEN
            FOR i := 1 TO count - 1 DO
                fifo[i] := fifo[i + 1];
            END_FOR
            fifo[count] := 0;
            count := count - 1;
        END_IF
    END_IF

    // push rising edge: add item if not full
    IF pushEn AND NOT prevPush THEN
        IF count < 8 THEN
            count := count + 1;
            fifo[count] := pushItem;
        END_IF
    END_IF

    // outputs
    full  := (count = 8);
    empty := (count = 0);
    head  := 0;
    IF NOT empty THEN
        head := fifo[1];
    END_IF

    // update edge detection history
    prevPush := pushEn;
    prevPop  := popEn;
END_FUNCTION_BLOCK

(* ---- self-hard-05.candidate_01.st ---- *)
FUNCTION_BLOCK FB
VAR_INPUT
    runRequest   : BOOL;
    flameOK      : BOOL;
    o2Valid      : BOOL;
    o2PV         : REAL;
    baseAir      : REAL;
    resetBtn     : BOOL;
END_VAR

VAR_OUTPUT
    fuelPermit   : BOOL;
    trimEnable   : BOOL;
    airTrim      : REAL;
    airCommand   : REAL;
    tripLatched  : BOOL;
    o2Fault      : BOOL;
END_VAR

VAR
    LatchTrip    : BOOL;      // internal latch for trip state
    prevResetBtn : BOOL;      // previous state of reset button for edge detection
END_VAR

// ---- Oxygen analyser fault detection ----
o2Fault := NOT o2Valid OR o2PV < 0.0 OR o2PV > 21.0;

// ---- Flame‑loss latch ----
// Set the latch the moment a flame loss occurs while the burner is requested to run
IF runRequest AND NOT flameOK THEN
    LatchTrip := TRUE;
END_IF

// Reset the latch only on the rising edge of the reset button when the burner is safely stopped
IF resetBtn AND NOT prevResetBtn AND NOT runRequest AND NOT flameOK THEN
    LatchTrip := FALSE;
END_IF

tripLatched := LatchTrip;

// ---- Fuel permit ----
fuelPermit := runRequest AND flameOK AND NOT LatchTrip;

// ---- Oxygen trim enable ----
trimEnable := fuelPermit AND NOT o2Fault;

// ---- Air trim bias ----
IF trimEnable THEN
    airTrim := 2.0 * (2.0 - o2PV);            // raw bias
    // clamp to ±10 %
    IF airTrim > 10.0 THEN
        airTrim := 10.0;
    END_IF;
    IF airTrim < -10.0 THEN
        airTrim := -10.0;
    END_IF;
ELSE
    airTrim := 0.0;
END_IF;

// ---- Air damper command ----
IF fuelPermit THEN
    airCommand := baseAir + airTrim;         // raw command
    // clamp final command to 0 % … 100 %
    IF airCommand > 100.0 THEN
        airCommand := 100.0;
    END_IF;
    IF airCommand < 0.0 THEN
        airCommand := 0.0;
    END_IF;
ELSE
    airCommand := 0.0;
END_IF;

// ---- Update edge‑detection variable ----
prevResetBtn := resetBtn;

END_FUNCTION_BLOCK
